ABB RAPID module: PrecProg.mod

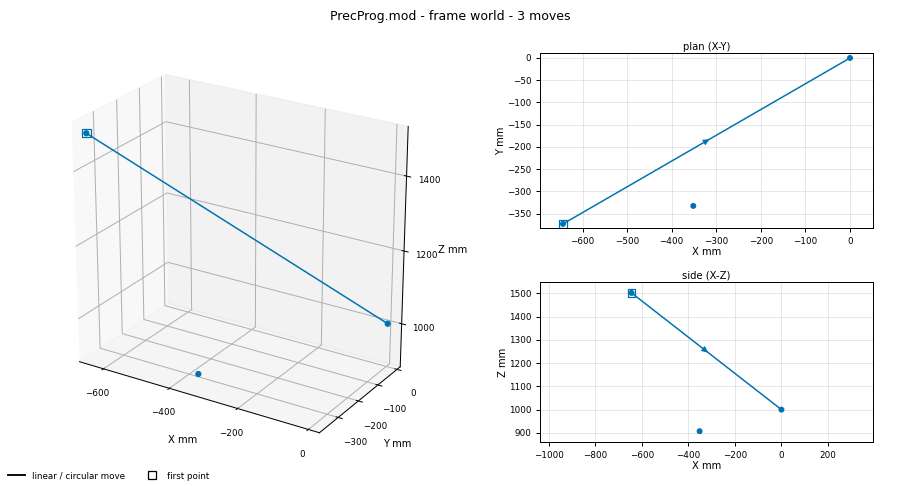
[picture p0: tool path of PrecProg.mod in frame world, 3 of 6 moves have a stored position in this frame; points joined in program order, loops and branches not executed]
%%%
  VERSION:1
  LANGUAGE:ENGLISH
%%%
MODULE MOD_PrecProg

    ! -------------------------------
    ! Define customized variables here
    ! ...

	! Tool variables:
	PERS tooldata ToolP := [TRUE,[[0.125,-0.375,123.457],[0.92304245,-0.38469811,-0.00000034,0.00000081]],[1,[0,0,20],[1,0,0,0],0,0,0.005]];

	! Reference variables:
	PERS wobjdata FrameP := [FALSE, TRUE, "", [[0,0,0],[1,0,0,0]],[[0.000,-0.001,1000.000],[0.70709693,0.70710235,-0.00232357,0.00384708]]];

	PROC Main()
		ConfJ \On;
		ConfL \Off;
		! Program generated by RoboDK v6.0.7 for ABB IRBT 2005 Standard 2.8m on XX/XX/XXXX 18:00:00
		! Using nominal kinematics.
		MoveAbsJ [[12.345600,0.000000,0.000000,0.000000,0.000000,0.000000],[9E+09,9E+09,9E+09,9E+09,9E+09,9E+09]],v500,z1,ToolP \WObj:=FrameP;
		MoveL [[-640.585,506.981,371.534],[0.37535171,0.28421100,0.85462317,-0.21898501],[0,0,0,0],[9E+09,9E+09,9E+09,9E+09,9E+09,9E+09]],v500,z1,ToolP \WObj:=FrameP;
		MoveL [[0.500,-0.500,0.250],[0.00000000,1.00000000,0.00004363,0.00004363],[0,0,0,0],[9E+09,9E+09,9E+09,9E+09,9E+09,9E+09]],v500,z1,ToolP \WObj:=FrameP;
		MoveAbsJ [[-12.345400,0.000000,0.000000,0.000000,0.000000,0.000000],[9E+09,9E+09,9E+09,9E+09,9E+09,9E+09]],v500,z1,ToolP \WObj:=FrameP;
		MoveAbsJ [[-12.345400,0.000000,0.000000,0.000000,0.000000,0.000000],[9E+09,9E+09,9E+09,9E+09,9E+09,9E+09]],v500,z1,ToolP \WObj:=FrameP;
		WaitTime 0.002;
		WaitTime 1.000;
		MoveL [[-353.026,-90.135,331.702],[0.34432926,0.04805561,0.93307257,-0.09221494],[0,0,0,0],[9E+09,9E+09,9E+09,9E+09,9E+09,9E+09]],[66.67,500,5000,1000],z1,ToolP \WObj:=FrameP;
	ENDPROC

ENDMODULE
